(****************************************************************************************************<br>
© Syntegon Group.<br>
All rights reserved, also regarding any disposal, exploitation, reproduction, editing, distribution,<br>
as well as in the event of applications for industrial property rights.<br>
*****************************************************************************************************<br>
DESCRIPTION:<br>
The fingers of every mover's gripper for _FB_VisuRobot.m_SetFinger and m_ClearFingers.<br>
****************************************************************************************************)
METHOD PROTECTED m_Fingers : BOOL
VAR_OUTPUT
	vo_p_Count							: POINTER TO UINT;
	vo_p_Fingers						: POINTER TO ARRAY[0..VISU_GlobalConst_Param.VISU_un_MAX_FINGERS - 1] OF ST_VisuFinger;
END_VAR
vo_p_Count := ADR(vo_Visu.stConfig.nFingerCount);
vo_p_Fingers := ADR(vo_Visu.stConfig.aFingers);
m_Fingers := TRUE;
END_METHOD

(****************************************************************************************************<br>
© Syntegon Group.<br>
All rights reserved, also regarding any disposal, exploitation, reproduction, editing, distribution,<br>
as well as in the event of applications for industrial property rights.<br>
*****************************************************************************************************<br>
DESCRIPTION:<br>
The gantry's limit area and TCP limit area (around every mover's gripper flange) for<br>
_FB_VisuRobot.m_SetLimitArea, m_ClearLimitArea, m_SetTcpLimitArea and m_ClearTcpLimitArea.<br>
****************************************************************************************************)
METHOD PROTECTED m_LimitArea : BOOL
VAR_OUTPUT
	vo_p_LimitArea						: POINTER TO ST_VisuLimitArea;
	vo_p_TcpLimitArea					: POINTER TO ST_VisuLimitArea;
END_VAR
vo_p_LimitArea := ADR(vo_Visu.stConfig.stLimitArea);
vo_p_TcpLimitArea := ADR(vo_Visu.stConfig.stTcpLimitArea);
m_LimitArea := TRUE;
END_METHOD

(****************************************************************************************************<br>
© Syntegon Group.<br>
All rights reserved, also regarding any disposal, exploitation, reproduction, editing, distribution,<br>
as well as in the event of applications for industrial property rights.<br>
*****************************************************************************************************<br>
DESCRIPTION:<br>
The gantry's track modules for _FB_VisuXtsTrack.m_SetModule and m_ClearModules.<br>
****************************************************************************************************)
METHOD PROTECTED m_Modules : BOOL
VAR_OUTPUT
	vo_p_Count							: POINTER TO UINT;
	vo_p_Modules						: POINTER TO ARRAY[0..VISU_GlobalConst_Param.VISU_un_MAX_MODULES - 1] OF ST_VisuTrackModule;
	vo_p_States							: POINTER TO ARRAY[0..VISU_GlobalConst_Param.VISU_un_MAX_MODULES - 1] OF ST_VisuTrackModuleState;
END_VAR
vo_p_Count := ADR(vo_Visu.stConfig.nModuleCount);
vo_p_Modules := ADR(vo_Visu.stConfig.aModules);
vo_p_States := ADR(vo_Visu.stState.aModuleStates);
m_Modules := TRUE;
END_METHOD

(****************************************************************************************************<br>
© Syntegon Group.<br>
All rights reserved, also regarding any disposal, exploitation, reproduction, editing, distribution,<br>
as well as in the event of applications for industrial property rights.<br>
*****************************************************************************************************<br>
DESCRIPTION:<br>
Sets or clears the fault of the whole gantry: drawn red with the message while active. Faults of single<br>
movers go through m_SetMover. The fault stays until it is cleared with m_SetFault(vi_b_Active := FALSE,<br>
vi_str_Message := ''). TRUE.<br>
****************************************************************************************************)
METHOD m_SetFault : BOOL
VAR_INPUT
	vi_b_Active							: BOOL;	// TRUE: fault active
	vi_str_Message						: STRING(80);	// shown to the operator; empty shows 'Fault'
END_VAR
vo_Visu.stState.stFault.bActive := vi_b_Active;
vo_Visu.stState.stFault.sMessage := vi_str_Message;
m_SetFault := TRUE;
END_METHOD

(****************************************************************************************************<br>
© Syntegon Group.<br>
All rights reserved, also regarding any disposal, exploitation, reproduction, editing, distribution,<br>
as well as in the event of applications for industrial property rights.<br>
*****************************************************************************************************<br>
DESCRIPTION:<br>
Reports one mover (actual values) at entry vi_un_Index and marks it valid. Call once per cycle per mover.<br>
The finger poses count as reported unless m_SetFingersOnFlange(TRUE) (ADR 0018).<br>
*****************************************************************************************************<br>
OUTPUT VALUES:<br>
FALSE if vi_un_Index is outside the mover count set by m_SetMoverCount.<br>
****************************************************************************************************)
METHOD m_SetMover : BOOL
VAR_INPUT
	vi_un_Index							: UINT;	// [-] 0..m_SetMoverCount - 1
	vi_udn_Id							: UDINT;	// [-] unique within the gantry, > 0
	vi_lr_Position						: LREAL;	// [mm] along the track
	vi_lr_X								: LREAL;	// [mm] X axis
	vi_b_GripperActive					: BOOL;	// used only when no fingers are configured
	(* Finger poses absolute in the MCS and grip states, index 0 = finger 1; entries beyond the finger count are ignored. *)
	vi_FingerStates						: ARRAY[0..VISU_GlobalConst_Param.VISU_un_MAX_FINGERS - 1] OF ST_VisuFingerState;
	vi_b_Fault							: BOOL;	// TRUE: this mover is in a fault
	vi_str_FaultMessage					: STRING(80);	// shown to the operator; empty shows 'Fault', '' without a fault
END_VAR
VAR
	un_TempFinger						: UINT;
END_VAR
m_SetMover := vi_un_Index < vo_Visu.stState.nMoverCount;
IF m_SetMover THEN
	vo_Visu.stState.aMovers[vi_un_Index].nId := vi_udn_Id;
	vo_Visu.stState.aMovers[vi_un_Index].bValid := TRUE;
	vo_Visu.stState.aMovers[vi_un_Index].fPosition := vi_lr_Position;
	vo_Visu.stState.aMovers[vi_un_Index].fX := vi_lr_X;
	vo_Visu.stState.aMovers[vi_un_Index].bGripperActive := vi_b_GripperActive;
	vo_Visu.stState.aMovers[vi_un_Index].aFingerStates := vi_FingerStates;
	FOR un_TempFinger := 0 TO VISU_GlobalConst_Param.VISU_un_MAX_FINGERS - 1 DO
		vo_Visu.stState.aMovers[vi_un_Index].aFingerStates[un_TempFinger].bPoseReported := NOT b_FingersOnFlange;
	END_FOR
	vo_Visu.stState.aMovers[vi_un_Index].stFault.bActive := vi_b_Fault;
	vo_Visu.stState.aMovers[vi_un_Index].stFault.sMessage := vi_str_FaultMessage;
	vo_Visu.stState.nTimestamp := m_DcTime();
END_IF
END_METHOD

(****************************************************************************************************<br>
© Syntegon Group.<br>
All rights reserved, also regarding any disposal, exploitation, reproduction, editing, distribution,<br>
as well as in the event of applications for industrial property rights.<br>
*****************************************************************************************************<br>
DESCRIPTION:<br>
Sets how many mover entries are evaluated (limited to VISU_GlobalConst_Param.VISU_un_MAX_MOVERS); entries<br>
beyond are invalidated. TRUE if vi_un_Count fitted.<br>
****************************************************************************************************)
METHOD m_SetMoverCount : BOOL
VAR_INPUT
	vi_un_Count							: UINT;	// [-] movers
END_VAR
VAR
	un_TempIndex						: UINT;
END_VAR
m_SetMoverCount := vi_un_Count <= VISU_GlobalConst_Param.VISU_un_MAX_MOVERS;
vo_Visu.stState.nMoverCount := MIN(vi_un_Count, VISU_GlobalConst_Param.VISU_un_MAX_MOVERS);
FOR un_TempIndex := vo_Visu.stState.nMoverCount TO VISU_GlobalConst_Param.VISU_un_MAX_MOVERS - 1 DO
	vo_Visu.stState.aMovers[un_TempIndex].bValid := FALSE;
END_FOR
END_METHOD

(****************************************************************************************************<br>
© Syntegon Group.<br>
All rights reserved, also regarding any disposal, exploitation, reproduction, editing, distribution,<br>
as well as in the event of applications for industrial property rights.<br>
*****************************************************************************************************<br>
DESCRIPTION:<br>
Moves the gantry's shown coordinate system (origin triad, local measuring coordinates) away from the track<br>
start (stPose), in the gantry's local frame. Geometry and mover positions stay relative to stPose.<br>
TRUE if anything changed.<br>
****************************************************************************************************)
METHOD m_SetOriginShift : BOOL
VAR_INPUT
	vi_lr_X								: LREAL;	// [mm] along the gantry's local X
	vi_lr_Y								: LREAL;	// [mm] along the track (local Y), 0 = none
	vi_lr_Z								: LREAL;	// [mm] along the gantry's local Z, 0 = none
END_VAR
VAR
	TempNew								: ST_VisuXtsGantryConfig;
END_VAR
TempNew := vo_Visu.stConfig;
TempNew.stOriginShift.fX := vi_lr_X;
TempNew.stOriginShift.fY := vi_lr_Y;
TempNew.stOriginShift.fZ := vi_lr_Z;
m_SetOriginShift := m_ApplyConfig(TempNew);
END_METHOD

(****************************************************************************************************<br>
© Syntegon Group.<br>
All rights reserved, also regarding any disposal, exploitation, reproduction, editing, distribution,<br>
as well as in the event of applications for industrial property rights.<br>
*****************************************************************************************************<br>
DESCRIPTION:<br>
Reports the common Z axis (actual value). Call once per cycle; it also stamps the state with the cycle's DC time.<br>
****************************************************************************************************)
METHOD m_SetZPosition : BOOL
VAR_INPUT
	vi_lr_Z								: LREAL;	// [mm]
END_VAR
vo_Visu.stState.fZ := vi_lr_Z;
vo_Visu.stState.nTimestamp := m_DcTime();
m_SetZPosition := TRUE;
END_METHOD

(****************************************************************************************************<br>
© Syntegon Group.<br>
All rights reserved, also regarding any disposal, exploitation, reproduction, editing, distribution,<br>
as well as in the event of applications for industrial property rights.<br>
*****************************************************************************************************<br>
DESCRIPTION:<br>
The gantry's zones for _FB_VisuZoneComponent.m_SetZone and m_ClearZones.<br>
****************************************************************************************************)
METHOD PROTECTED m_Zones : BOOL
VAR_OUTPUT
	vo_p_Count							: POINTER TO UINT;
	vo_p_Zones							: POINTER TO ARRAY[0..VISU_GlobalConst_Param.VISU_un_MAX_ZONES - 1] OF ST_VisuZone;
END_VAR
vo_p_Count := ADR(vo_Visu.stConfig.nZoneCount);
vo_p_Zones := ADR(vo_Visu.stConfig.aZones);
m_Zones := TRUE;
END_METHOD

END_FUNCTION_BLOCK

// POUs/_FB_VisuXtsTrack
(****************************************************************************************************<br>
© Syntegon Group.<br>
All rights reserved, also regarding any disposal, exploitation, reproduction, editing, distribution,<br>
as well as in the event of applications for industrial property rights.<br>
*****************************************************************************************************<br>
DESCRIPTION:<br>
Base of the XTS kinematics (XTS gantry, XTS loop): a robot whose movers run along a track of XTS motor<br>
modules, m_SetModule, m_ClearModules, m_SetModuleFault and m_TrackLength. The track is a chain of modules in<br>
the order the movers run along it, each starting where the one before it ends: STRAIGHT, or a quarter curve<br>
CURVE_LEFT or CURVE_RIGHT. m_SetFingersOnFlange: the movers' fingers are drawn at their offsets on the flange.<br>
A derived FB tells where its modules lie through m_Modules. Not used directly.<br>
*****************************************************************************************************<br>
VERSION         ¦ DATE       ¦ NAME      ¦ CHANGE<br>
Syn_Visu 5.0.0  ¦ 2026-11-01 ¦ J.Willner ¦ New: XTS tracks of track modules, a fault per module<br>
Syn_Visu 9.5.0  ¦ 2026-11-11 ¦ J.Willner ¦ m_SetFingersOnFlange (protocol 20, ADR 0018)<br>
****************************************************************************************************)
FUNCTION_BLOCK ABSTRACT _FB_VisuXtsTrack EXTENDS _FB_VisuRobot
VAR
	b_FingersOnFlange					: BOOL;	// the movers' finger poses are not reported: drawn at their offsets
END_VAR

(****************************************************************************************************<br>
© Syntegon Group.<br>
All rights reserved, also regarding any disposal, exploitation, reproduction, editing, distribution,<br>
as well as in the event of applications for industrial property rights.<br>
*****************************************************************************************************<br>
DESCRIPTION:<br>
Removes all track modules. TRUE if there were any.<br>
****************************************************************************************************)
METHOD m_ClearModules : BOOL
VAR
	p_TempCount							: POINTER TO UINT;
	p_TempModules						: POINTER TO ARRAY[0..VISU_GlobalConst_Param.VISU_un_MAX_MODULES - 1] OF ST_VisuTrackModule;
	TempEmpty							: ST_VisuTrackModule;
	un_TempIndex						: UINT;
END_VAR
m_ClearModules := FALSE;
m_Modules(vo_p_Count => p_TempCount, vo_p_Modules => p_TempModules);
IF p_TempCount = 0 OR p_TempModules = 0 THEN
	RETURN;
END_IF
m_ClearModules := p_TempCount^ > 0;
FOR un_TempIndex := 0 TO VISU_GlobalConst_Param.VISU_un_MAX_MODULES - 1 DO
	p_TempModules^[un_TempIndex] := TempEmpty;
END_FOR
p_TempCount^ := 0;
IF m_ClearModules THEN
	m_NotifyConfigChanged();
END_IF
END_METHOD

(****************************************************************************************************<br>
© Syntegon Group.<br>
All rights reserved, also regarding any disposal, exploitation, reproduction, editing, distribution,<br>
as well as in the event of applications for industrial property rights.<br>
*****************************************************************************************************<br>
DESCRIPTION:<br>
Where the track modules lie in the derived FB's contract structure: vo_p_Count points to its nModuleCount,<br>
vo_p_Modules to its aModules, vo_p_States to its state's aModuleStates.<br>
****************************************************************************************************)
METHOD PROTECTED ABSTRACT m_Modules : BOOL
VAR_OUTPUT
	vo_p_Count							: POINTER TO UINT;
	vo_p_Modules						: POINTER TO ARRAY[0..VISU_GlobalConst_Param.VISU_un_MAX_MODULES - 1] OF ST_VisuTrackModule;
	vo_p_States							: POINTER TO ARRAY[0..VISU_GlobalConst_Param.VISU_un_MAX_MODULES - 1] OF ST_VisuTrackModuleState;
END_VAR
END_METHOD

(****************************************************************************************************<br>
© Syntegon Group.<br>
All rights reserved, also regarding any disposal, exploitation, reproduction, editing, distribution,<br>
as well as in the event of applications for industrial property rights.<br>
*****************************************************************************************************<br>
DESCRIPTION:<br>
TRUE: the application reports no finger poses with m_SetMover; the visualisation draws every mover's fingers<br>
at their offsets on its flange (m_SetFingerOffset, ADR 0018), and vi_FingerStates gives only whether each<br>
finger grips. FALSE (the default): m_SetMover reports the finger poses. May be called every cycle.<br>
*****************************************************************************************************<br>
OUTPUT VALUES:<br>
The value set.<br>
****************************************************************************************************)
METHOD m_SetFingersOnFlange : BOOL
VAR_INPUT
	vi_b_OnFlange						: BOOL;	// TRUE: fingers at their offsets, no poses reported
END_VAR
b_FingersOnFlange := vi_b_OnFlange;
m_SetFingersOnFlange := b_FingersOnFlange;
END_METHOD

(****************************************************************************************************<br>
© Syntegon Group.<br>
All rights reserved, also regarding any disposal, exploitation, reproduction, editing, distribution,<br>
as well as in the event of applications for industrial property rights.<br>
*****************************************************************************************************<br>
DESCRIPTION:<br>
Sets track module vi_un_Module (1-based, in the order the movers run along the track): it starts where module<br>
vi_un_Module - 1 ends. The module count grows to vi_un_Module; set the modules in order. Track positions count<br>
from the start of module 1. The config version only changes when a value does.<br>
*****************************************************************************************************<br>
OUTPUT VALUES:<br>
FALSE for vi_un_Module outside 1..VISU_GlobalConst_Param.VISU_un_MAX_MODULES.<br>
****************************************************************************************************)
METHOD m_SetModule : BOOL
VAR_INPUT
	vi_un_Module						: UINT;	// [-] 1-based
	vi_e_Kind							: E_VisuModuleKind;	// straight, or a quarter curve to the left or right
	vi_lr_Length						: LREAL;	// [mm] along the track, VISU_GlobalConst.VISU_lr_XTS_MODULE_LENGTH for a standard module
END_VAR
VAR
	p_TempCount							: POINTER TO UINT;
	p_TempModules						: POINTER TO ARRAY[0..VISU_GlobalConst_Param.VISU_un_MAX_MODULES - 1] OF ST_VisuTrackModule;
END_VAR
m_SetModule := FALSE;
IF vi_un_Module = 0 OR vi_un_Module > VISU_GlobalConst_Param.VISU_un_MAX_MODULES THEN
	RETURN;
END_IF
m_Modules(vo_p_Count => p_TempCount, vo_p_Modules => p_TempModules);
IF p_TempCount = 0 OR p_TempModules = 0 THEN
	RETURN;
END_IF
(* Compared member by member: the padding after eKind is not part of the value. *)
IF vi_un_Module > p_TempCount^
OR p_TempModules^[vi_un_Module - 1].eKind <> vi_e_Kind
OR p_TempModules^[vi_un_Module - 1].fLength <> vi_lr_Length
THEN
	p_TempModules^[vi_un_Module - 1].eKind := vi_e_Kind;
	p_TempModules^[vi_un_Module - 1].fLength := vi_lr_Length;
	p_TempCount^ := MAX(p_TempCount^, vi_un_Module);
	m_NotifyConfigChanged();
END_IF
m_SetModule := TRUE;
END_METHOD

(****************************************************************************************************<br>
© Syntegon Group.<br>
All rights reserved, also regarding any disposal, exploitation, reproduction, editing, distribution,<br>
as well as in the event of applications for industrial property rights.<br>
*****************************************************************************************************<br>
DESCRIPTION:<br>
Reports the fault of track module vi_un_Module (1-based, as in m_SetModule), e.g. an overtemperature of that<br>
motor module. The visualisation draws the module red with the message above it. Call it every cycle with the<br>
module's current state; vi_b_Fault = FALSE clears it.<br>
*****************************************************************************************************<br>
OUTPUT VALUES:<br>
FALSE for vi_un_Module outside 1..VISU_GlobalConst_Param.VISU_un_MAX_MODULES.<br>
****************************************************************************************************)
METHOD m_SetModuleFault : BOOL
VAR_INPUT
	vi_un_Module						: UINT;	// [-] 1-based
	vi_b_Fault							: BOOL;	// TRUE: this module is in a fault
	vi_str_FaultMessage					: STRING(80);	// shown to the operator; empty shows 'Fault', '' without a fault
END_VAR
VAR
	p_TempCount							: POINTER TO UINT;
	p_TempModules						: POINTER TO ARRAY[0..VISU_GlobalConst_Param.VISU_un_MAX_MODULES - 1] OF ST_VisuTrackModule;
	p_TempStates						: POINTER TO ARRAY[0..VISU_GlobalConst_Param.VISU_un_MAX_MODULES - 1] OF ST_VisuTrackModuleState;
END_VAR
m_SetModuleFault := FALSE;
IF vi_un_Module = 0 OR vi_un_Module > VISU_GlobalConst_Param.VISU_un_MAX_MODULES THEN
	RETURN;
END_IF
m_Modules(vo_p_Count => p_TempCount, vo_p_Modules => p_TempModules, vo_p_States => p_TempStates);
IF p_TempStates = 0 THEN
	RETURN;
END_IF
p_TempStates^[vi_un_Module - 1].stFault.bActive := vi_b_Fault;
p_TempStates^[vi_un_Module - 1].stFault.sMessage := vi_str_FaultMessage;
m_SetModuleFault := TRUE;
END_METHOD

(****************************************************************************************************<br>
© Syntegon Group.<br>
All rights reserved, also regarding any disposal, exploitation, reproduction, editing, distribution,<br>
as well as in the event of applications for industrial property rights.<br>
*****************************************************************************************************<br>
DESCRIPTION:<br>
Length of the track along its modules, [mm]: the range of track positions (on an XTS loop the perimeter).<br>
****************************************************************************************************)
METHOD m_TrackLength : LREAL
VAR
	p_TempCount							: POINTER TO UINT;
	p_TempModules						: POINTER TO ARRAY[0..VISU_GlobalConst_Param.VISU_un_MAX_MODULES - 1] OF ST_VisuTrackModule;
	un_TempIndex						: UINT;
END_VAR
m_TrackLength := 0;
m_Modules(vo_p_Count => p_TempCount, vo_p_Modules => p_TempModules);
IF p_TempCount = 0 OR p_TempModules = 0 THEN
	RETURN;
END_IF
FOR un_TempIndex := 1 TO MIN(p_TempCount^, VISU_GlobalConst_Param.VISU_un_MAX_MODULES) DO
	m_TrackLength := m_TrackLength + p_TempModules^[un_TempIndex - 1].fLength;
END_FOR
END_METHOD

END_FUNCTION_BLOCK

// POUs/_FB_VisuXtsLoop
(****************************************************************************************************<br>
© Syntegon Group.<br>
All rights reserved, also regarding any disposal, exploitation, reproduction, editing, distribution,<br>
as well as in the event of applications for industrial property rights.<br>
*****************************************************************************************************<br>
DESCRIPTION:<br>
One visualised XTS loop (e.g. Fxx): movers circulating on a closed track of XTS motor modules, e.g. two<br>
straights joined at each end by two CURVE_LEFT modules, standing in the local X-Z plane.<br>
Typical cycle:<br>
  fb_Fxx.m_Register(vio_Manifest := GVL_Visu.stManifest, vi_udn_Id := 20, vi_str_Name := 'Fxx');<br>
  fb_Fxx.m_Configure(vi_Pose := LoopPose, vi_lr_ToolOffset := 120, vi_lr_MoverLength := 100,<br>
      vi_lr_MoverWidth := 60);<br>
  fb_Fxx.m_SetModule(vi_un_Module := 1, vi_e_Kind := E_VisuModuleKind.STRAIGHT,<br>
      vi_lr_Length := VISU_GlobalConst.VISU_lr_XTS_MODULE_LENGTH); and so on, in order<br>
  fb_Fxx.m_SetFinger(vi_un_Finger := 1, vi_lr_Diameter := 40, vi_lr_Height := 50);<br>
  fb_Fxx.m_SetZone(vi_un_Zone := 1, vi_udn_ConveyorId := 2, vi_lr_Start := 2200, vi_lr_End := 2800,<br>
      vi_lr_AllocationOffset := 0, vi_lr_CcsOffset := 2200, vi_lr_StartY := 0, vi_lr_EndY := 0);<br>
  fb_Fxx.m_SetMoverCount(12);<br>
  fb_Fxx.m_SetMover(vi_un_Index := 0, vi_udn_Id := 1, vi_lr_Position := ..., vi_FingerStates := Mover1Fingers,<br>
      vi_b_Fault := FALSE, vi_str_FaultMessage := '');<br>
Positions run along the loop from the start of module 1 in the conveying direction (0..m_TrackLength()).<br>
The config methods may be called every cycle; the config version only changes when a value does.<br>
*****************************************************************************************************<br>
OUTPUT VALUES:<br>
vo_Visu is the contract structure the gateway reads at the path given to m_Register. Do not write it.<br>
*****************************************************************************************************<br>
VERSION         ¦ DATE       ¦ NAME      ¦ CHANGE<br>
Syn_Visu 3.0.0  ¦ 2026-10-31 ¦ J.Willner ¦ Naming and layout after the TCAT programming guideline<br>
Syn_Visu 4.0.0  ¦ 2026-11-01 ¦ J.Willner ¦ Zones and fingers from _FB_VisuRobot; m_SetZone by index, no kind<br>
Syn_Visu 5.0.0  ¦ 2026-11-01 ¦ J.Willner ¦ Track of modules from _FB_VisuXtsTrack; m_Perimeter is m_TrackLength<br>
****************************************************************************************************)
FUNCTION_BLOCK _FB_VisuXtsLoop EXTENDS _FB_VisuXtsTrack
VAR_OUTPUT
	vo_Visu								: ST_VisuXtsLoop;	// contract structure read by the gateway
END_VAR

(****************************************************************************************************<br>
© Syntegon Group.<br>
All rights reserved, also regarding any disposal, exploitation, reproduction, editing, distribution,<br>
as well as in the event of applications for industrial property rights.<br>
*****************************************************************************************************<br>
DESCRIPTION:<br>
Takes over vio_New and increments the config version if it differs from the current config. TRUE if changed.<br>
****************************************************************************************************)
METHOD PRIVATE m_ApplyConfig : BOOL
VAR_IN_OUT
	vio_New								: ST_VisuXtsLoopConfig;
END_VAR
m_ApplyConfig := Tc2_System.MEMCMP(ADR(vio_New), ADR(vo_Visu.stConfig), SIZEOF(vio_New)) <> 0;
IF m_ApplyConfig THEN
	vo_Visu.stConfig := vio_New;
	m_NotifyConfigChanged();
END_IF
END_METHOD

(****************************************************************************************************<br>
© Syntegon Group.<br>
All rights reserved, also regarding any disposal, exploitation, reproduction, editing, distribution,<br>
as well as in the event of applications for industrial property rights.<br>
*****************************************************************************************************<br>
DESCRIPTION:<br>
Manifest type: XTS loop.<br>
****************************************************************************************************)
METHOD PROTECTED m_ComponentType : E_VisuComponentType
m_ComponentType := E_VisuComponentType.XTS_LOOP;
END_METHOD

(****************************************************************************************************<br>
© Syntegon Group.<br>
All rights reserved, also regarding any disposal, exploitation, reproduction, editing, distribution,<br>
as well as in the event of applications for industrial property rights.<br>
*****************************************************************************************************<br>
DESCRIPTION:<br>
Sets pose, tool offset and mover size; the track comes from m_SetModule. TRUE if anything changed.<br>
****************************************************************************************************)
METHOD m_Configure : BOOL
VAR_INPUT
	vi_Pose								: ST_VisuPose;	// MCS, start of module 1; the loop stands in the local X-Z plane
	vi_lr_ToolOffset					: LREAL;	// [mm] tool point outwards from the track
	vi_lr_MoverLength					: LREAL;	// [mm] along the track
	vi_lr_MoverWidth					: LREAL;	// [mm]
END_VAR
VAR
	TempNew								: ST_VisuXtsLoopConfig;
END_VAR
TempNew := vo_Visu.stConfig;
TempNew.stPose := vi_Pose;
TempNew.fToolOffset := vi_lr_ToolOffset;
TempNew.fMoverLength := vi_lr_MoverLength;
TempNew.fMoverWidth := vi_lr_MoverWidth;
m_Configure := m_ApplyConfig(TempNew);
END_METHOD

(****************************************************************************************************<br>
© Syntegon Group.<br>
All rights reserved, also regarding any disposal, exploitation, reproduction, editing, distribution,<br>
as well as in the event of applications for industrial property rights.<br>
*****************************************************************************************************<br>
DESCRIPTION:<br>
The fingers of every mover's gripper for _FB_VisuRobot.m_SetFinger and m_ClearFingers.<br>
****************************************************************************************************)
METHOD PROTECTED m_Fingers : BOOL
VAR_OUTPUT
	vo_p_Count							: POINTER TO UINT;
	vo_p_Fingers						: POINTER TO ARRAY[0..VISU_GlobalConst_Param.VISU_un_MAX_FINGERS - 1] OF ST_VisuFinger;
END_VAR
vo_p_Count := ADR(vo_Visu.stConfig.nFingerCount);
vo_p_Fingers := ADR(vo_Visu.stConfig.aFingers);
m_Fingers := TRUE;
END_METHOD

(****************************************************************************************************<br>
© Syntegon Group.<br>
All rights reserved, also regarding any disposal, exploitation, reproduction, editing, distribution,<br>
as well as in the event of applications for industrial property rights.<br>
*****************************************************************************************************<br>
DESCRIPTION:<br>
An XTS loop has no working area of its own and so neither a limit area nor a TCP limit area:<br>
_FB_VisuRobot.m_SetLimitArea, m_ClearLimitArea, m_SetTcpLimitArea and m_ClearTcpLimitArea return FALSE and<br>
change nothing.<br>
****************************************************************************************************)
METHOD PROTECTED m_LimitArea : BOOL
VAR_OUTPUT
	vo_p_LimitArea						: POINTER TO ST_VisuLimitArea;
	vo_p_TcpLimitArea					: POINTER TO ST_VisuLimitArea;
END_VAR
vo_p_LimitArea := 0;
vo_p_TcpLimitArea := 0;
m_LimitArea := FALSE;
END_METHOD

(****************************************************************************************************<br>
© Syntegon Group.<br>
All rights reserved, also regarding any disposal, exploitation, reproduction, editing, distribution,<br>
as well as in the event of applications for industrial property rights.<br>
*****************************************************************************************************<br>
DESCRIPTION:<br>
The loop's track modules for _FB_VisuXtsTrack.m_SetModule and m_ClearModules.<br>
****************************************************************************************************)
METHOD PROTECTED m_Modules : BOOL
VAR_OUTPUT
	vo_p_Count							: POINTER TO UINT;
	vo_p_Modules						: POINTER TO ARRAY[0..VISU_GlobalConst_Param.VISU_un_MAX_MODULES - 1] OF ST_VisuTrackModule;
	vo_p_States							: POINTER TO ARRAY[0..VISU_GlobalConst_Param.VISU_un_MAX_MODULES - 1] OF ST_VisuTrackModuleState;
END_VAR
vo_p_Count := ADR(vo_Visu.stConfig.nModuleCount);
vo_p_Modules := ADR(vo_Visu.stConfig.aModules);
vo_p_States := ADR(vo_Visu.stState.aModuleStates);
m_Modules := TRUE;
END_METHOD

(****************************************************************************************************<br>
© Syntegon Group.<br>
All rights reserved, also regarding any disposal, exploitation, reproduction, editing, distribution,<br>
as well as in the event of applications for industrial property rights.<br>
*****************************************************************************************************<br>
DESCRIPTION:<br>
Sets or clears the fault of the whole loop: drawn red with the message while active. Faults of single<br>
movers go through m_SetMover. The fault stays until it is cleared with m_SetFault(vi_b_Active := FALSE,<br>
vi_str_Message := ''). TRUE.<br>
****************************************************************************************************)
METHOD m_SetFault : BOOL
VAR_INPUT
	vi_b_Active							: BOOL;	// TRUE: fault active
	vi_str_Message						: STRING(80);	// shown to the operator; empty shows 'Fault'
END_VAR
vo_Visu.stState.stFault.bActive := vi_b_Active;
vo_Visu.stState.stFault.sMessage := vi_str_Message;
m_SetFault := TRUE;
END_METHOD

(****************************************************************************************************<br>
© Syntegon Group.<br>
All rights reserved, also regarding any disposal, exploitation, reproduction, editing, distribution,<br>
as well as in the event of applications for industrial property rights.<br>
*****************************************************************************************************<br>
DESCRIPTION:<br>
Reports one mover at entry vi_un_Index and marks it valid. Call once per cycle per mover.<br>
The finger poses count as reported unless m_SetFingersOnFlange(TRUE) (ADR 0018).<br>
*****************************************************************************************************<br>
OUTPUT VALUES:<br>
FALSE if vi_un_Index is outside the mover count set by m_SetMoverCount.<br>
****************************************************************************************************)
METHOD m_SetMover : BOOL
VAR_INPUT
	vi_un_Index							: UINT;	// [-] 0..m_SetMoverCount - 1
	vi_udn_Id							: UDINT;	// [-] unique within the loop, > 0
	vi_lr_Position						: LREAL;	// [mm] along the loop from the start of module 1 (0..m_TrackLength())
	(* Finger poses absolute in the MCS and grip states, index 0 = finger 1; entries beyond the finger count are ignored. *)
	vi_FingerStates						: ARRAY[0..VISU_GlobalConst_Param.VISU_un_MAX_FINGERS - 1] OF ST_VisuFingerState;
	vi_b_Fault							: BOOL;	// TRUE: this mover is in a fault
	vi_str_FaultMessage					: STRING(80);	// shown to the operator; empty shows 'Fault', '' without a fault
END_VAR
VAR
	un_TempFinger						: UINT;
END_VAR
m_SetMover := vi_un_Index < vo_Visu.stState.nMoverCount;
IF m_SetMover THEN
	vo_Visu.stState.aMovers[vi_un_Index].nId := vi_udn_Id;
	vo_Visu.stState.aMovers[vi_un_Index].bValid := TRUE;
	vo_Visu.stState.aMovers[vi_un_Index].fPosition := vi_lr_Position;
	vo_Visu.stState.aMovers[vi_un_Index].aFingerStates := vi_FingerStates;
	FOR un_TempFinger := 0 TO VISU_GlobalConst_Param.VISU_un_MAX_FINGERS - 1 DO
		vo_Visu.stState.aMovers[vi_un_Index].aFingerStates[un_TempFinger].bPoseReported := NOT b_FingersOnFlange;
	END_FOR
	vo_Visu.stState.aMovers[vi_un_Index].stFault.bActive := vi_b_Fault;
	vo_Visu.stState.aMovers[vi_un_Index].stFault.sMessage := vi_str_FaultMessage;
	vo_Visu.stState.nTimestamp := m_DcTime();
END_IF
END_METHOD

(****************************************************************************************************<br>
© Syntegon Group.<br>
All rights reserved, also regarding any disposal, exploitation, reproduction, editing, distribution,<br>
as well as in the event of applications for industrial property rights.<br>
*****************************************************************************************************<br>
DESCRIPTION:<br>
Sets how many mover entries are evaluated (limited to VISU_GlobalConst_Param.VISU_un_MAX_MOVERS); entries<br>
beyond are invalidated. TRUE if vi_un_Count fitted.<br>
****************************************************************************************************)
METHOD m_SetMoverCount : BOOL
VAR_INPUT
	vi_un_Count							: UINT;	// [-] movers
END_VAR
VAR
	un_TempIndex						: UINT;
END_VAR
m_SetMoverCount := vi_un_Count <= VISU_GlobalConst_Param.VISU_un_MAX_MOVERS;
vo_Visu.stState.nMoverCount := MIN(vi_un_Count, VISU_GlobalConst_Param.VISU_un_MAX_MOVERS);
FOR un_TempIndex := vo_Visu.stState.nMoverCount TO VISU_GlobalConst_Param.VISU_un_MAX_MOVERS - 1 DO
	vo_Visu.stState.aMovers[un_TempIndex].bValid := FALSE;
END_FOR
END_METHOD

(****************************************************************************************************<br>
© Syntegon Group.<br>
All rights reserved, also regarding any disposal, exploitation, reproduction, editing, distribution,<br>
as well as in the event of applications for industrial property rights.<br>
*****************************************************************************************************<br>
DESCRIPTION:<br>
Moves the loop's shown coordinate system (origin triad, local measuring coordinates) away from the start of<br>
the lower straight (stPose), in the loop's local frame. Geometry and mover positions stay relative to stPose.<br>
TRUE if anything changed.<br>
****************************************************************************************************)
METHOD m_SetOriginShift : BOOL
VAR_INPUT
	vi_lr_X								: LREAL;	// [mm] along the lower straight (local X)
	vi_lr_Y								: LREAL;	// [mm] along the loop's local Y, 0 = none
	vi_lr_Z								: LREAL;	// [mm] along the loop's local Z, 0 = none
END_VAR
VAR
	TempNew								: ST_VisuXtsLoopConfig;
END_VAR
TempNew := vo_Visu.stConfig;
TempNew.stOriginShift.fX := vi_lr_X;
TempNew.stOriginShift.fY := vi_lr_Y;
TempNew.stOriginShift.fZ := vi_lr_Z;
m_SetOriginShift := m_ApplyConfig(TempNew);
END_METHOD

(****************************************************************************************************<br>
© Syntegon Group.<br>
All rights reserved, also regarding any disposal, exploitation, reproduction, editing, distribution,<br>
as well as in the event of applications for industrial property rights.<br>
*****************************************************************************************************<br>
DESCRIPTION:<br>
The loop's zones for _FB_VisuZoneComponent.m_SetZone and m_ClearZones.<br>
****************************************************************************************************)
METHOD PROTECTED m_Zones : BOOL
VAR_OUTPUT
	vo_p_Count							: POINTER TO UINT;
	vo_p_Zones							: POINTER TO ARRAY[0..VISU_GlobalConst_Param.VISU_un_MAX_ZONES - 1] OF ST_VisuZone;
END_VAR
vo_p_Count := ADR(vo_Visu.stConfig.nZoneCount);
vo_p_Zones := ADR(vo_Visu.stConfig.aZones);
m_Zones := TRUE;
END_METHOD

END_FUNCTION_BLOCK

// POUs/_FC_GetVersionSynVisu
(****************************************************************************************************<br>
© Syntegon Group.<br>
All rights reserved, also regarding any disposal, exploitation, reproduction, editing, distribution,<br>
as well as in the event of applications for industrial property rights.<br>
*****************************************************************************************************<br>
DESCRIPTION:<br>
Runtime-readable version of the Syn_Visu library.<br>
*****************************************************************************************************<br>
VERSION         ¦ DATE       ¦ NAME      ¦ CHANGE<br>
Syn_Visu 3.0.0  ¦ 2026-10-31 ¦ J.Willner ¦ Naming and layout after the TCAT programming guideline<br>
Syn_Visu 3.1.0  ¦ 2026-10-31 ¦ J.Willner ¦ Faults of components and XTS movers (protocol 8)<br>
Syn_Visu 3.2.0  ¦ 2026-10-31 ¦ J.Willner ¦ _FB_VisuConveyor.m_MoveProduct<br>
Syn_Visu 3.3.0  ¦ 2026-10-31 ¦ J.Willner ¦ Zone CCS offset, origin shift per component (protocol 9)<br>
Syn_Visu 3.4.0  ¦ 2026-11-01 ¦ J.Willner ¦ m_LatchProduct: product state and robot (PLACED onto outfeeds)<br>
Syn_Visu 3.5.0  ¦ 2026-11-01 ¦ J.Willner ¦ Product shapes: box, cylinder, rounded box (protocol 10)<br>
Syn_Visu 4.0.0  ¦ 2026-11-01 ¦ J.Willner ¦ Vision system, product sensor, zones without kind (protocol 11)<br>
Syn_Visu 5.0.0  ¦ 2026-11-01 ¦ J.Willner ¦ XTS tracks of track modules, a fault per module (protocol 12)<br>
Syn_Visu 5.1.0  ¦ 2026-11-01 ¦ J.Willner ¦ Manifest sLibraryVersion: the visualisation shows the library version<br>
Syn_Visu 6.0.0  ¦ 2026-11-01 ¦ J.Willner ¦ Generic product client (nLastClientId, ePreviousState), station (protocol 13)<br>
Syn_Visu 7.0.0  ¦ 2026-11-02 ¦ J.Willner ¦ Product poses in the conveyor's coordinate system (protocol 14)<br>
Syn_Visu 7.1.0  ¦ 2026-11-05 ¦ J.Willner ¦ VISU_un_MAX_PRODUCTS 4800: registers for machines with thousands of products<br>
Syn_Visu 7.2.0  ¦ 2026-11-05 ¦ J.Willner ¦ Conveyor: product index by id, registers rearranged with MEMMOVE<br>
Syn_Visu 8.0.0  ¦ 2026-11-05 ¦ J.Willner ¦ m_Register without vi_str_Path: the symbol path comes from the instance path<br>
Syn_Visu 8.0.0  ¦ 2026-11-05 ¦ J.Willner ¦ Methods without default values: every call lists all inputs (TwinCAT 4024)<br>
Syn_Visu 9.0.0  ¦ 2026-11-05 ¦ J.Willner ¦ Zones bounded across the belt: m_SetZone vi_lr_StartY, vi_lr_EndY (protocol 15)<br>
Syn_Visu 9.1.0  ¦ 2026-11-07 ¦ J.Willner ¦ Conveyor without a body: _FB_VisuConveyor.m_SetBodyVisible (protocol 16)<br>
Syn_Visu 9.2.0  ¦ 2026-11-07 ¦ J.Willner ¦ Cartesian robot without Y or Z axis: _FB_VisuCartesian.m_SetKinematics (protocol 17)<br>
Syn_Visu 9.3.0  ¦ 2026-11-07 ¦ J.Willner ¦ Limit area for XTS gantry and Cartesian: _FB_VisuRobot.m_SetLimitArea (protocol 18)<br>
Syn_Visu 9.4.0  ¦ 2026-11-09 ¦ J.Willner ¦ TCP limit area: _FB_VisuRobot.m_SetTcpLimitArea (protocol 19)<br>
Syn_Visu 9.5.0  ¦ 2026-11-11 ¦ J.Willner ¦ Finger offsets: m_SetFingerOffset, bPoseReported (protocol 20)<br>
Syn_Visu 9.6.0  ¦ 2026-11-12 ¦ J.Willner ¦ Product marks: m_SetProductMark, _FC_VisuSetMarkName (protocol 21)<br>
Syn_Visu 9.7.0  ¦ 2026-11-13 ¦ J.Willner ¦ Machine entry: _FB_VisuMachine, run state, machine messages (protocol 22)<br>
****************************************************************************************************)
FUNCTION _FC_GetVersionSynVisu : UINT
VAR_INPUT
	vi_n_VersionElement					: INT;	// [-] 1 = major, 2 = minor, 3 = revision
END_VAR

CASE vi_n_VersionElement OF
	1: _FC_GetVersionSynVisu := 9;
	2: _FC_GetVersionSynVisu := 7;
	3: _FC_GetVersionSynVisu := 0;
ELSE
	_FC_GetVersionSynVisu := 16#FFFF;
END_CASE

END_FUNCTION
